// TIA Portal V20 export
Screen "Pop-up_Device"  395x540
  ScreenItem "Text field TG Status" at 1,0 size 393x47  Type=HmiTextBox
  ScreenItem "Cancel Mode" at 316,3 size 76x42  Type=HmiButton
  ScreenItem "Background_1" at 0,37 size 368x32  Type=HmiRectangle
  ScreenItem "Text field TG1 Status_22" at 9,41 size 126x21  Type=HmiTextBox
  ScreenItem "Text field TG1 Status_1" at 191,43 size 78x21  Type=HmiTextBox
  ScreenItem "Rectangle TG1" at 1,74 size 367x40  Type=HmiRectangle
  ScreenItem "Textfeld_2" at 191,85 size 245x20  Type=HmiTextBox
  ScreenItem "Rectangle TG1_1" at 1,113 size 367x40  Type=HmiRectangle
  ScreenItem "Rectangle TG1_2" at 1,156 size 367x40  Type=HmiRectangle
  ScreenItem "Rectangle TG1_3" at 1,238 size 367x40  Type=HmiRectangle
  ScreenItem "Rectangle TG1_4" at 1,197 size 367x40  Type=HmiRectangle
  ScreenItem "Textfeld_13" at 191,126 size 275x20  Type=HmiTextBox
  ScreenItem "Textfeld_14" at 191,167 size 275x20  Type=HmiTextBox
  ScreenItem "Textfeld_15" at 191,208 size 110x20  Type=HmiTextBox
  ScreenItem "Textfeld_21" at 191,249 size 275x20  Type=HmiTextBox
  ScreenItem "Background_2" at 0,0 size 368x32  Type=HmiRectangle
  ScreenItem "Text field TG1 Status_2" at 142,7 size 126x21  Type=HmiTextBox
  ScreenItem "Text_Symbol_PN-DEV_OK" at 11,83 size 24x20  Type=HmiTextBox
  ScreenItem "Textfeld_1" at 43,83 size 19x20  Type=HmiTextBox
  ScreenItem "Text_Symbol_PN-DEV_OK_1" at 11,124 size 24x20  Type=HmiTextBox
  ScreenItem "Textfeld_4" at 43,124 size 19x20  Type=HmiTextBox
  ScreenItem "Text_Symbol_PN-DEV_OK_2" at 11,165 size 24x20  Type=HmiTextBox
  ScreenItem "Textfeld_5" at 43,165 size 19x20  Type=HmiTextBox
  ScreenItem "Text_Symbol_PN-DEV_OK_3" at 11,206 size 24x20  Type=HmiTextBox
  ScreenItem "Textfeld_6" at 43,206 size 19x20  Type=HmiTextBox
  ScreenItem "Text_Symbol_PN-DEV_OK_4" at 11,247 size 24x20  Type=HmiTextBox
  ScreenItem "Textfeld_8" at 43,247 size 44x20  Type=HmiTextBox
  ScreenItem "Rectangle TG1_5" at 1,279 size 367x40  Type=HmiRectangle
  ScreenItem "Rectangle TG1_10" at 1,320 size 367x40  Type=HmiRectangle
  ScreenItem "Line_1" at 114,74 size 3x285  Type=HmiLine
  ScreenItem "Text_Symbol_PN-DEV_OK_5" at 11,286 size 24x20  Type=HmiTextBox
  ScreenItem "Textfeld_10" at 43,286 size 44x20  Type=HmiTextBox
  ScreenItem "Text_Symbol_PN-DEV_OK_6" at 11,332 size 24x20  Type=HmiTextBox
  ScreenItem "Textfeld_17" at 43,332 size 44x20  Type=HmiTextBox
  ScreenItem "Textfeld_20" at 191,290 size 275x20  Type=HmiTextBox
  ScreenItem "Textfeld_22" at 191,332 size 275x20  Type=HmiTextBox
  ScreenItem "Background_3" at 0,37 size 368x32  Type=HmiRectangle
  ScreenItem "Text field TG1 Status_3" at 9,41 size 126x21  Type=HmiTextBox
  ScreenItem "Text field TG1 Status_4" at 191,43 size 78x21  Type=HmiTextBox
  ScreenItem "Rectangle TG1_8" at 1,74 size 367x40  Type=HmiRectangle
  ScreenItem "Background_4" at 0,0 size 368x32  Type=HmiRectangle
  ScreenItem "Text field TG1 Status_5" at 112,7 size 126x21  Type=HmiTextBox
  ScreenItem "Text_Symbol_PN-DEV_OK_13" at 11,83 size 24x20  Type=HmiTextBox
  ScreenItem "Textfeld_18" at 43,83 size 19x20  Type=HmiTextBox
  ScreenItem "Line_2" at 114,74 size 0x39  Type=HmiLine
  ScreenItem "Textfeld_19" at 183,83 size 245x20  Type=HmiTextBox
